FUNCTION_BLOCK basicGeradorGenerico (* Logica unica do grupo gerador (DEIF AGC 150): valores, estado do QTA, modo e alarmes *)
  (* Standard: 61499-2 *)
  (* Version 1.1, 15/10/2026, Hidryco, Hidryco, 1.1: comandos basicos (automatico, semiautomatico, partir, parar, reconhecer alarmes do AGC) nas palavras 5 e 6. 1.0: AGC 150 (GEN) por Modbus TCP FC04, tabela DEIF rev. S; so supervisao *)
  PACKAGE Hidryco.HidrycoLib;
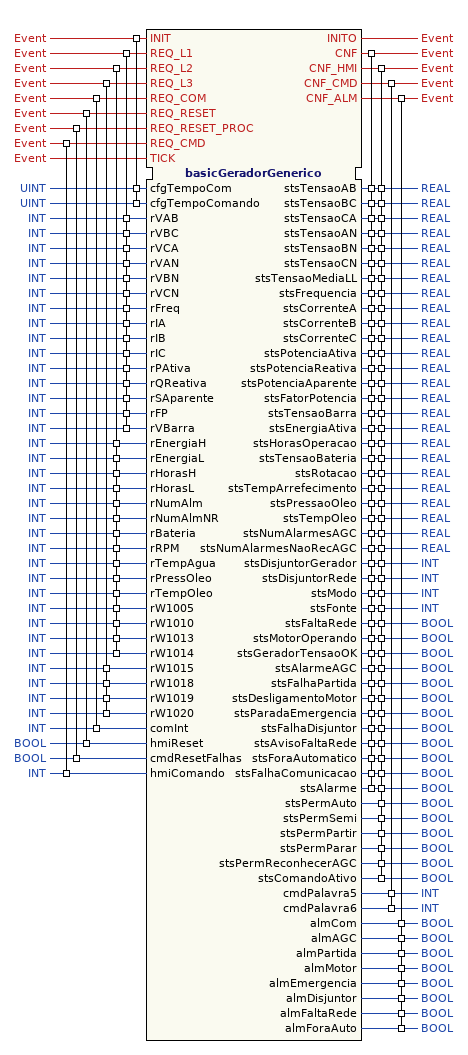
  EVENT_INPUT
    INIT WITH cfgTempoCom, cfgTempoComando; (* Inicializacao *)
    REQ_L1 WITH rVAB, rVBC, rVCA, rVAN, rVBN, rVCN, rFreq, rIA, rIB, rIC, rPAtiva, rQReativa, rSAparente, rFP, rVBarra; (* Leitura 1 (grandezas eletricas) *)
    REQ_L2 WITH rEnergiaH, rEnergiaL, rHorasH, rHorasL, rNumAlm, rNumAlmNR, rBateria, rRPM, rTempAgua, rPressOleo, rTempOleo, rW1005, rW1010, rW1013, rW1014; (* Leitura 2 (contadores, motor, alarmes) *)
    REQ_L3 WITH rW1015, rW1018, rW1019, rW1020; (* Leitura 3 (estado e modos) *)
    REQ_COM WITH comInt; (* Comunicacao *)
    REQ_RESET WITH hmiReset; (* Reconhecimento pela IHM *)
    REQ_RESET_PROC WITH cmdResetFalhas; (* Reconhecimento pelo processo *)
    REQ_CMD WITH hmiComando; (* Comando da IHM para o AGC *)
    TICK; (* Base de tempo de 1 s (E_CYCLE) *)
  END_EVENT
  EVENT_OUTPUT
    INITO; (* Inicializacao concluida *)
    CNF WITH stsTensaoAB, stsTensaoBC, stsTensaoCA, stsTensaoAN, stsTensaoBN, stsTensaoCN, stsTensaoMediaLL, stsFrequencia, stsCorrenteA, stsCorrenteB, stsCorrenteC, stsPotenciaAtiva, stsPotenciaReativa, stsPotenciaAparente, stsFatorPotencia, stsTensaoBarra, stsEnergiaAtiva, stsHorasOperacao, stsTensaoBateria, stsRotacao, stsTempArrefecimento, stsPressaoOleo, stsTempOleo, stsNumAlarmesAGC, stsNumAlarmesNaoRecAGC, stsDisjuntorGerador, stsDisjuntorRede, stsModo, stsFonte, stsFaltaRede, stsMotorOperando, stsGeradorTensaoOK, stsAlarmeAGC, stsFalhaPartida, stsDesligamentoMotor, stsParadaEmergencia, stsFalhaDisjuntor, stsAvisoFaltaRede, stsForaAutomatico, stsFalhaComunicacao, stsAlarme; (* Valores e estados (na mudanca) *)
    CNF_HMI WITH stsTensaoAB, stsTensaoBC, stsTensaoCA, stsTensaoAN, stsTensaoBN, stsTensaoCN, stsTensaoMediaLL, stsFrequencia, stsCorrenteA, stsCorrenteB, stsCorrenteC, stsPotenciaAtiva, stsPotenciaReativa, stsPotenciaAparente, stsFatorPotencia, stsTensaoBarra, stsEnergiaAtiva, stsHorasOperacao, stsTensaoBateria, stsRotacao, stsTempArrefecimento, stsPressaoOleo, stsTempOleo, stsNumAlarmesAGC, stsNumAlarmesNaoRecAGC, stsDisjuntorGerador, stsDisjuntorRede, stsModo, stsFonte, stsFaltaRede, stsMotorOperando, stsGeradorTensaoOK, stsAlarmeAGC, stsFalhaPartida, stsDesligamentoMotor, stsParadaEmergencia, stsFalhaDisjuntor, stsAvisoFaltaRede, stsForaAutomatico, stsFalhaComunicacao, stsAlarme, stsPermAuto, stsPermSemi, stsPermPartir, stsPermParar, stsPermReconhecerAGC, stsComandoAtivo; (* Status para a IHM (na mudanca) *)
    CNF_CMD WITH cmdPalavra5, cmdPalavra6; (* Palavras de comando do AGC (na mudanca) *)
    CNF_ALM WITH almCom, almAGC, almPartida, almMotor, almEmergencia, almDisjuntor, almFaltaRede, almForaAuto; (* Alarmes para os ALARM_BIT (na mudanca) *)
  END_EVENT
  VAR_INPUT
    cfgTempoCom : UINT := 10; (* Tempo (s) sem comunicacao com o AGC 150 para confirmar a falha *)
    cfgTempoComando : UINT := 2; (* Tempo (s) que a palavra de comando fica escrita no AGC *)
    rVAB : INT; (* Tensao do gerador L1-L2 (V) *)
    rVBC : INT; (* Tensao do gerador L2-L3 (V) *)
    rVCA : INT; (* Tensao do gerador L3-L1 (V) *)
    rVAN : INT; (* Tensao do gerador L1-N (V) *)
    rVBN : INT; (* Tensao do gerador L2-N (V) *)
    rVCN : INT; (* Tensao do gerador L3-N (V) *)
    rFreq : INT; (* Frequencia do gerador L1 (0,01 Hz) *)
    rIA : INT; (* Corrente do gerador L1 (A) *)
    rIB : INT; (* Corrente do gerador L2 (A) *)
    rIC : INT; (* Corrente do gerador L3 (A) *)
    rPAtiva : INT; (* Potencia ativa do gerador (kW) *)
    rQReativa : INT; (* Potencia reativa do gerador (kVAr) *)
    rSAparente : INT; (* Potencia aparente do gerador (kVA) *)
    rFP : INT; (* Fator de potencia do gerador (0,01) *)
    rVBarra : INT; (* Tensao do lado B (barramento/rede) L1-L2 (V) *)
    rEnergiaH : INT; (* Energia ativa exportada total - palavra alta (INT32 ABCD, kWh) *)
    rEnergiaL : INT; (* Energia ativa exportada total - palavra baixa *)
    rHorasH : INT; (* Horas de funcionamento absolutas - palavra alta (INT32 ABCD, h) *)
    rHorasL : INT; (* Horas de funcionamento absolutas - palavra baixa *)
    rNumAlm : INT; (* Numero de alarmes ativos no AGC *)
    rNumAlmNR : INT; (* Numero de alarmes nao reconhecidos no AGC *)
    rBateria : INT; (* Tensao de alimentacao DC (bateria), term. 1-2 (0,1 V) *)
    rRPM : INT; (* Rotacao do motor - ECU (rpm) *)
    rTempAgua : INT; (* Temperatura do liquido de arrefecimento - ECU (0,1 C) *)
    rPressOleo : INT; (* Pressao do oleo - ECU (0,01 bar) *)
    rTempOleo : INT; (* Temperatura do oleo - ECU (0,1 C) *)
    rW1005 : INT; (* Alarmes de disjuntor e sincronismo (bits) *)
    rW1010 : INT; (* Alarmes de entradas digitais (bit 12 = parada de emergencia) *)
    rW1013 : INT; (* Alarmes do motor (bits: 9/10 sobrevelocidade, 11 falha de arranque, 15 falha de partida) *)
    rW1014 : INT; (* Alarmes do motor (bit 0 = falha de parada) *)
    rW1015 : INT; (* Alarmes diversos (bit 12 = fora do automatico) *)
    rW1018 : INT; (* Estado da planta (bits: 0 falta de rede, 1 MB ON, 4 GB ON, 6 motor em operacao, 8 Hz/V OK, 11 GB OFF, 12 MB OFF) *)
    rW1019 : INT; (* Modos (bits: 0 bloqueio, 1 manual, 2 semi-auto, 3 auto, 4 teste) *)
    rW1020 : INT; (* Alarmes da ECU (bit 2 = shutdown / alarme vermelho) *)
    comInt : INT; (* connStatusInt do MODBUSGENTCPS (1 = online) *)
    hmiReset : BOOL; (* IHM: reconhecimento *)
    cmdResetFalhas : BOOL; (* Processo: reconhecimento (com E_RESET_FALHAS) *)
    hmiComando : INT; (* IHM: comando para o AGC (1 automatico, 2 semiautomatico, 3 partir, 4 parar, 5 reconhecer alarmes do AGC) *)
  END_VAR
  VAR_OUTPUT
    stsTensaoAB : REAL; (* Tensao A-B (V) *)
    stsTensaoBC : REAL; (* Tensao B-C (V) *)
    stsTensaoCA : REAL; (* Tensao C-A (V) *)
    stsTensaoAN : REAL; (* Tensao A-N (V) *)
    stsTensaoBN : REAL; (* Tensao B-N (V) *)
    stsTensaoCN : REAL; (* Tensao C-N (V) *)
    stsTensaoMediaLL : REAL; (* Tensao media fase-fase (V) *)
    stsFrequencia : REAL; (* Frequencia (Hz) *)
    stsCorrenteA : REAL; (* Corrente fase A (A) *)
    stsCorrenteB : REAL; (* Corrente fase B (A) *)
    stsCorrenteC : REAL; (* Corrente fase C (A) *)
    stsPotenciaAtiva : REAL; (* Potencia ativa (kW) *)
    stsPotenciaReativa : REAL; (* Potencia reativa (kVAr) *)
    stsPotenciaAparente : REAL; (* Potencia aparente (kVA) *)
    stsFatorPotencia : REAL; (* Fator de potencia *)
    stsTensaoBarra : REAL; (* Tensao do lado B (barramento/rede) L1-L2 (V) *)
    stsEnergiaAtiva : REAL; (* Energia ativa exportada (kWh) *)
    stsHorasOperacao : REAL; (* Horas de funcionamento (h) *)
    stsTensaoBateria : REAL; (* Tensao da bateria (V) *)
    stsRotacao : REAL; (* Rotacao do motor (rpm) *)
    stsTempArrefecimento : REAL; (* Temperatura do liquido de arrefecimento (°C) *)
    stsPressaoOleo : REAL; (* Pressao do oleo (bar) *)
    stsTempOleo : REAL; (* Temperatura do oleo (°C) *)
    stsNumAlarmesAGC : REAL; (* Alarmes ativos no AGC *)
    stsNumAlarmesNaoRecAGC : REAL; (* Alarmes nao reconhecidos no AGC *)
    stsDisjuntorGerador : INT; (* Disjuntor do gerador (GB): 0 indefinido/sem comunicacao, 1 aberto, 2 fechado *)
    stsDisjuntorRede : INT; (* Disjuntor de rede (MB): 0 indefinido/sem comunicacao, 1 aberto, 2 fechado *)
    stsModo : INT; (* Modo do AGC: 0 indefinido, 1 automatico, 2 semi-automatico, 3 manual, 4 bloqueio, 5 teste *)
    stsFonte : INT; (* Fonte da saida do QTA: 0 sem fonte, 1 rede, 2 gerador, 3 indefinida (sem comunicacao) *)
    stsFaltaRede : BOOL; (* Falta de rede (AMF) *)
    stsMotorOperando : BOOL; (* Motor em operacao *)
    stsGeradorTensaoOK : BOOL; (* Tensao e frequencia do gerador OK *)
    stsAlarmeAGC : BOOL; (* Alarme ativo no controlador do gerador (AGC 150) *)
    stsFalhaPartida : BOOL; (* Falha na partida do gerador *)
    stsDesligamentoMotor : BOOL; (* Desligamento do motor (ECU ou sobrevelocidade) *)
    stsParadaEmergencia : BOOL; (* Parada de emergência do gerador acionada *)
    stsFalhaDisjuntor : BOOL; (* Falha de disjuntor no QTA (gerador ou rede) *)
    stsAvisoFaltaRede : BOOL; (* Falta de rede no QTA *)
    stsForaAutomatico : BOOL; (* Gerador fora do modo automático *)
    stsFalhaComunicacao : BOOL; (* Falha de comunicacao com o AGC 150 *)
    stsAlarme : BOOL; (* Algum alarme do gerador *)
    stsPermAuto : BOOL; (* IHM: comando Auto permitido *)
    stsPermSemi : BOOL; (* IHM: comando Semi permitido *)
    stsPermPartir : BOOL; (* IHM: comando Partir permitido *)
    stsPermParar : BOOL; (* IHM: comando Parar permitido *)
    stsPermReconhecerAGC : BOOL; (* IHM: comando ReconhecerAGC permitido *)
    stsComandoAtivo : BOOL; (* Comando sendo enviado ao AGC *)
    cmdPalavra5 : INT; (* Palavra de comando 5 do AGC (holding register 5) *)
    cmdPalavra6 : INT; (* Palavra de comando 6 do AGC (holding register 6) *)
    almCom : BOOL; (* ALARM_BIT falha de comunicacao *)
    almAGC : BOOL; (* ALARM_BIT Alarme ativo no controlador do gerador (AGC 150) *)
    almPartida : BOOL; (* ALARM_BIT Falha na partida do gerador *)
    almMotor : BOOL; (* ALARM_BIT Desligamento do motor (ECU ou sobrevelocidade) *)
    almEmergencia : BOOL; (* ALARM_BIT Parada de emergência do gerador acionada *)
    almDisjuntor : BOOL; (* ALARM_BIT Falha de disjuntor no QTA (gerador ou rede) *)
    almFaltaRede : BOOL; (* ALARM_BIT Falta de rede no QTA *)
    almForaAuto : BOOL; (* ALARM_BIT Gerador fora do modo automático *)
  END_VAR
  VAR
    initDone : BOOL;
    initPass : BOOL;
    bComRecebida : BOOL; (* Ja houve leitura do connStatusInt *)
    bValido : BOOL; (* AGC comunicando: valores validos *)
    uSegCom : UDINT;
    w05 : WORD;
    w10 : WORD;
    w13 : WORD;
    w18 : WORD;
    w19 : WORD;
    w20 : WORD;
    bGBon : BOOL;
    bGBoff : BOOL;
    bMBon : BOOL;
    bMBoff : BOOL;
    bMudou : BOOL;
    wSts : DWORD;
    oldSts : DWORD := 16#FFFFFFFF;
    wAlm : WORD;
    oldAlm : WORD := 16#FFFF;
    iOld : INT;
    uCmd : UINT; (* Segundos restantes do pulso de comando *)
    wPerm : WORD;
    oldPerm : WORD := 16#FFFF;
    o_stsTensaoAB : REAL := -1.0;
    o_stsTensaoBC : REAL := -1.0;
    o_stsTensaoCA : REAL := -1.0;
    o_stsTensaoAN : REAL := -1.0;
    o_stsTensaoBN : REAL := -1.0;
    o_stsTensaoCN : REAL := -1.0;
    o_stsTensaoMediaLL : REAL := -1.0;
    o_stsFrequencia : REAL := -1.0;
    o_stsCorrenteA : REAL := -1.0;
    o_stsCorrenteB : REAL := -1.0;
    o_stsCorrenteC : REAL := -1.0;
    o_stsPotenciaAtiva : REAL := -1.0;
    o_stsPotenciaReativa : REAL := -1.0;
    o_stsPotenciaAparente : REAL := -1.0;
    o_stsFatorPotencia : REAL := -1.0;
    o_stsTensaoBarra : REAL := -1.0;
    o_stsEnergiaAtiva : REAL := -1.0;
    o_stsHorasOperacao : REAL := -1.0;
    o_stsTensaoBateria : REAL := -1.0;
    o_stsRotacao : REAL := -1.0;
    o_stsTempArrefecimento : REAL := -1.0;
    o_stsPressaoOleo : REAL := -1.0;
    o_stsTempOleo : REAL := -1.0;
    o_stsNumAlarmesAGC : REAL := -1.0;
    o_stsNumAlarmesNaoRecAGC : REAL := -1.0;
    o_stsDisjuntorGerador : INT := -1;
    o_stsDisjuntorRede : INT := -1;
    o_stsModo : INT := -1;
    o_stsFonte : INT := -1;
  END_VAR
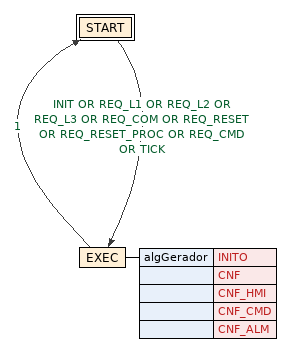
  EC_STATES
    START; (* Estado inicial *)
    EXEC : algGerador -> INITO, -> CNF, -> CNF_HMI, -> CNF_CMD, -> CNF_ALM; (* Executa a logica; o algoritmo decide quais eventos saem *)
  END_STATES
  EC_TRANSITIONS
    START TO EXEC := INIT OR REQ_L1 OR REQ_L2 OR REQ_L3 OR REQ_COM OR REQ_RESET OR REQ_RESET_PROC OR REQ_CMD OR TICK;
    EXEC TO START := 1;
  END_TRANSITIONS
  ALGORITHM algGerador IN ST: (* Logica completa do gerador (um unico algoritmo) *)
(* =====================================================================
   basicGeradorGenerico v1.0 - grupo gerador com controlador DEIF AGC 150
   (aplicacao GEN: QTA com disjuntor do gerador GB e de rede MB)
   Registradores de entrada (FC04) da tabela DEIF "AGC 150 Modbus server
   tables" rev. S (software 1.19). v1.1: comandos basicos nas palavras de
   comando 5 e 6 (pulso de cfgTempoComando s; depois as palavras voltam a 0).
   Padrao das bibliotecas Schneider: eventos de saida desligados no inicio e
   ligados so na mudanca; tempos contados pelo TICK de 1 s (E_CYCLE do CAT).
   - escalas da tabela: frequencia e FP 0,01; bateria, temperaturas 0,1;
     pressao do oleo 0,01 bar; energia e horas INT32 (ABCD, palavra alta 1o);
   - falha de comunicacao: connStatusInt <> 1 por cfgTempoCom s; com a
     falha os estados ficam indefinidos e os demais alarmes suprimidos;
   - alarmes seguem o AGC (nao memorizados aqui): o reconhecimento na IHM
     reconhece os ALARM_BIT; os alarmes do AGC sao reconhecidos no AGC.
   ===================================================================== *)

INITO   := FALSE;
CNF     := FALSE;
CNF_HMI := FALSE;
CNF_CMD := FALSE;
CNF_ALM := FALSE;

IF REQ_COM THEN
    bComRecebida := TRUE;
END_IF;
IF INIT THEN
    initDone := TRUE;
    initPass := TRUE;
    INITO    := TRUE;
END_IF;
IF NOT initDone THEN
    RETURN;
END_IF;

(* ---- 1. Comunicacao ---- *)
IF comInt <> 1 THEN
    IF TICK AND uSegCom < UINT_TO_UDINT(cfgTempoCom) THEN
        uSegCom := uSegCom + 1;
    END_IF;
ELSE
    uSegCom := 0;
END_IF;
stsFalhaComunicacao := comInt <> 1 AND uSegCom >= UINT_TO_UDINT(cfgTempoCom);
bValido := bComRecebida AND comInt = 1;

(* ---- 2. Valores (ficam congelados sem comunicacao) ---- *)
stsTensaoAB := INT_TO_REAL(rVAB);
stsTensaoBC := INT_TO_REAL(rVBC);
stsTensaoCA := INT_TO_REAL(rVCA);
stsTensaoAN := INT_TO_REAL(rVAN);
stsTensaoBN := INT_TO_REAL(rVBN);
stsTensaoCN := INT_TO_REAL(rVCN);
stsTensaoMediaLL := (INT_TO_REAL(rVAB) + INT_TO_REAL(rVBC) + INT_TO_REAL(rVCA)) / 3.0;
stsFrequencia := INT_TO_REAL(rFreq) / 100.0;
stsCorrenteA := INT_TO_REAL(rIA);
stsCorrenteB := INT_TO_REAL(rIB);
stsCorrenteC := INT_TO_REAL(rIC);
stsPotenciaAtiva := INT_TO_REAL(rPAtiva);
stsPotenciaReativa := INT_TO_REAL(rQReativa);
stsPotenciaAparente := INT_TO_REAL(rSAparente);
stsFatorPotencia := INT_TO_REAL(rFP) / 100.0;
stsTensaoBarra := INT_TO_REAL(rVBarra);
stsEnergiaAtiva := DINT_TO_REAL(DWORD_TO_DINT(SHL(WORD_TO_DWORD(INT_TO_WORD(rEnergiaH)), 16) OR WORD_TO_DWORD(INT_TO_WORD(rEnergiaL))));
stsHorasOperacao := DINT_TO_REAL(DWORD_TO_DINT(SHL(WORD_TO_DWORD(INT_TO_WORD(rHorasH)), 16) OR WORD_TO_DWORD(INT_TO_WORD(rHorasL))));
stsTensaoBateria := INT_TO_REAL(rBateria) / 10.0;
stsRotacao := INT_TO_REAL(rRPM);
stsTempArrefecimento := INT_TO_REAL(rTempAgua) / 10.0;
stsPressaoOleo := INT_TO_REAL(rPressOleo) / 100.0;
stsTempOleo := INT_TO_REAL(rTempOleo) / 10.0;
stsNumAlarmesAGC := INT_TO_REAL(rNumAlm);
stsNumAlarmesNaoRecAGC := INT_TO_REAL(rNumAlmNR);

(* ---- 3. Palavras de estado e alarme ---- *)
w05 := INT_TO_WORD(rW1005);
w10 := INT_TO_WORD(rW1010);
w13 := INT_TO_WORD(rW1013);
w18 := INT_TO_WORD(rW1018);
w19 := INT_TO_WORD(rW1019);
w20 := INT_TO_WORD(rW1020);
bGBon  := (w18 AND 16#0010) <> 16#0000;
bGBoff := (w18 AND 16#0800) <> 16#0000;
bMBon  := (w18 AND 16#0002) <> 16#0000;
bMBoff := (w18 AND 16#1000) <> 16#0000;

stsFaltaRede := bValido AND ((w18 AND 16#0001) <> 16#0000);
stsMotorOperando := bValido AND ((w18 AND 16#0040) <> 16#0000);
stsGeradorTensaoOK := bValido AND ((w18 AND 16#0100) <> 16#0000);

(* disjuntores: 2 fechado, 1 aberto, 0 indefinido (transicao ou sem comunicacao) *)
IF NOT bValido THEN
    stsDisjuntorGerador := 0;
    stsDisjuntorRede := 0;
ELSE
    IF bGBon AND NOT bGBoff THEN stsDisjuntorGerador := 2;
    ELSIF bGBoff AND NOT bGBon THEN stsDisjuntorGerador := 1;
    ELSE stsDisjuntorGerador := 0;
    END_IF;
    IF bMBon AND NOT bMBoff THEN stsDisjuntorRede := 2;
    ELSIF bMBoff AND NOT bMBon THEN stsDisjuntorRede := 1;
    ELSE stsDisjuntorRede := 0;
    END_IF;
END_IF;

(* modo: teste > bloqueio > manual > semi > auto *)
IF NOT bValido THEN stsModo := 0;
ELSIF (w19 AND 16#0010) <> 16#0000 THEN stsModo := 5;
ELSIF (w19 AND 16#0001) <> 16#0000 THEN stsModo := 4;
ELSIF (w19 AND 16#0002) <> 16#0000 THEN stsModo := 3;
ELSIF (w19 AND 16#0004) <> 16#0000 THEN stsModo := 2;
ELSIF (w19 AND 16#0008) <> 16#0000 THEN stsModo := 1;
ELSE stsModo := 0;
END_IF;

(* fonte da saida do QTA *)
IF NOT bValido THEN stsFonte := 3;
ELSIF stsDisjuntorGerador = 2 THEN stsFonte := 2;
ELSIF stsDisjuntorRede = 2 THEN stsFonte := 1;
ELSE stsFonte := 0;
END_IF;

(* ---- 4. Alarmes (seguem o AGC; so com comunicacao) ---- *)
stsAlarmeAGC := bValido AND (rNumAlm > 0);
stsFalhaPartida := bValido AND ((w13 AND 16#8800) <> 16#0000);
stsDesligamentoMotor := bValido AND (((w20 AND 16#0004) <> 16#0000) OR ((w13 AND 16#0600) <> 16#0000));
stsParadaEmergencia := bValido AND ((w10 AND 16#1000) <> 16#0000);
stsFalhaDisjuntor := bValido AND ((w05 AND 16#03F0) <> 16#0000);
stsAvisoFaltaRede := bValido AND ((w18 AND 16#0001) <> 16#0000);
stsForaAutomatico := bValido AND ((w19 AND 16#0008) = 16#0000);

almCom := stsFalhaComunicacao;
almAGC := stsAlarmeAGC;
almPartida := stsFalhaPartida;
almMotor := stsDesligamentoMotor;
almEmergencia := stsParadaEmergencia;
almDisjuntor := stsFalhaDisjuntor;
almFaltaRede := stsAvisoFaltaRede;
almForaAuto := stsForaAutomatico;
stsAlarme := almCom OR almAGC OR almPartida OR almMotor OR almEmergencia OR almDisjuntor OR almFaltaRede OR almForaAuto;

(* ---- 5. Comandos basicos (IHM) nas palavras 5 e 6 do AGC ---- *)
stsPermAuto := bValido AND stsModo <> 1;
stsPermSemi := bValido AND stsModo <> 2;
stsPermPartir := bValido AND stsModo = 2 AND NOT stsMotorOperando;
stsPermParar := bValido AND stsModo = 2 AND stsMotorOperando;
stsPermReconhecerAGC := bValido;
IF REQ_CMD AND uCmd = 0 THEN
    IF hmiComando = 1 AND stsPermAuto THEN
        cmdPalavra6 := 8193; cmdPalavra5 := 0;
        uCmd := cfgTempoComando + 1;
        CNF_CMD := TRUE;
    ELSIF hmiComando = 2 AND stsPermSemi THEN
        cmdPalavra6 := 16385; cmdPalavra5 := 0;
        uCmd := cfgTempoComando + 1;
        CNF_CMD := TRUE;
    ELSIF hmiComando = 3 AND stsPermPartir THEN
        cmdPalavra5 := 3; cmdPalavra6 := 0;
        uCmd := cfgTempoComando + 1;
        CNF_CMD := TRUE;
    ELSIF hmiComando = 4 AND stsPermParar THEN
        cmdPalavra5 := 17; cmdPalavra6 := 0;
        uCmd := cfgTempoComando + 1;
        CNF_CMD := TRUE;
    ELSIF hmiComando = 5 AND stsPermReconhecerAGC THEN
        cmdPalavra5 := 1025; cmdPalavra6 := 0;
        uCmd := cfgTempoComando + 1;
        CNF_CMD := TRUE;
    END_IF;
END_IF;
IF TICK AND uCmd > 0 THEN
    uCmd := uCmd - 1;
    IF uCmd = 0 THEN
        cmdPalavra5 := 0;
        cmdPalavra6 := 0;
        CNF_CMD := TRUE;
    END_IF;
END_IF;
IF NOT bValido AND uCmd > 0 THEN
    uCmd := 0;
    cmdPalavra5 := 0;
    cmdPalavra6 := 0;
    CNF_CMD := TRUE;
END_IF;
stsComandoAtivo := uCmd > 0;
wPerm := 0;
IF stsPermAuto THEN wPerm := wPerm OR 16#0001; END_IF;
IF stsPermSemi THEN wPerm := wPerm OR 16#0002; END_IF;
IF stsPermPartir THEN wPerm := wPerm OR 16#0004; END_IF;
IF stsPermParar THEN wPerm := wPerm OR 16#0008; END_IF;
IF stsPermReconhecerAGC THEN wPerm := wPerm OR 16#0010; END_IF;
IF stsComandoAtivo THEN wPerm := wPerm OR 16#0020; END_IF;

(* ---- 6. Eventos so na mudanca ---- *)
bMudou := FALSE;
IF stsTensaoAB <> o_stsTensaoAB THEN bMudou := TRUE; o_stsTensaoAB := stsTensaoAB; END_IF;
IF stsTensaoBC <> o_stsTensaoBC THEN bMudou := TRUE; o_stsTensaoBC := stsTensaoBC; END_IF;
IF stsTensaoCA <> o_stsTensaoCA THEN bMudou := TRUE; o_stsTensaoCA := stsTensaoCA; END_IF;
IF stsTensaoAN <> o_stsTensaoAN THEN bMudou := TRUE; o_stsTensaoAN := stsTensaoAN; END_IF;
IF stsTensaoBN <> o_stsTensaoBN THEN bMudou := TRUE; o_stsTensaoBN := stsTensaoBN; END_IF;
IF stsTensaoCN <> o_stsTensaoCN THEN bMudou := TRUE; o_stsTensaoCN := stsTensaoCN; END_IF;
IF stsTensaoMediaLL <> o_stsTensaoMediaLL THEN bMudou := TRUE; o_stsTensaoMediaLL := stsTensaoMediaLL; END_IF;
IF stsFrequencia <> o_stsFrequencia THEN bMudou := TRUE; o_stsFrequencia := stsFrequencia; END_IF;
IF stsCorrenteA <> o_stsCorrenteA THEN bMudou := TRUE; o_stsCorrenteA := stsCorrenteA; END_IF;
IF stsCorrenteB <> o_stsCorrenteB THEN bMudou := TRUE; o_stsCorrenteB := stsCorrenteB; END_IF;
IF stsCorrenteC <> o_stsCorrenteC THEN bMudou := TRUE; o_stsCorrenteC := stsCorrenteC; END_IF;
IF stsPotenciaAtiva <> o_stsPotenciaAtiva THEN bMudou := TRUE; o_stsPotenciaAtiva := stsPotenciaAtiva; END_IF;
IF stsPotenciaReativa <> o_stsPotenciaReativa THEN bMudou := TRUE; o_stsPotenciaReativa := stsPotenciaReativa; END_IF;
IF stsPotenciaAparente <> o_stsPotenciaAparente THEN bMudou := TRUE; o_stsPotenciaAparente := stsPotenciaAparente; END_IF;
IF stsFatorPotencia <> o_stsFatorPotencia THEN bMudou := TRUE; o_stsFatorPotencia := stsFatorPotencia; END_IF;
IF stsTensaoBarra <> o_stsTensaoBarra THEN bMudou := TRUE; o_stsTensaoBarra := stsTensaoBarra; END_IF;
IF stsEnergiaAtiva <> o_stsEnergiaAtiva THEN bMudou := TRUE; o_stsEnergiaAtiva := stsEnergiaAtiva; END_IF;
IF stsHorasOperacao <> o_stsHorasOperacao THEN bMudou := TRUE; o_stsHorasOperacao := stsHorasOperacao; END_IF;
IF stsTensaoBateria <> o_stsTensaoBateria THEN bMudou := TRUE; o_stsTensaoBateria := stsTensaoBateria; END_IF;
IF stsRotacao <> o_stsRotacao THEN bMudou := TRUE; o_stsRotacao := stsRotacao; END_IF;
IF stsTempArrefecimento <> o_stsTempArrefecimento THEN bMudou := TRUE; o_stsTempArrefecimento := stsTempArrefecimento; END_IF;
IF stsPressaoOleo <> o_stsPressaoOleo THEN bMudou := TRUE; o_stsPressaoOleo := stsPressaoOleo; END_IF;
IF stsTempOleo <> o_stsTempOleo THEN bMudou := TRUE; o_stsTempOleo := stsTempOleo; END_IF;
IF stsNumAlarmesAGC <> o_stsNumAlarmesAGC THEN bMudou := TRUE; o_stsNumAlarmesAGC := stsNumAlarmesAGC; END_IF;
IF stsNumAlarmesNaoRecAGC <> o_stsNumAlarmesNaoRecAGC THEN bMudou := TRUE; o_stsNumAlarmesNaoRecAGC := stsNumAlarmesNaoRecAGC; END_IF;
IF stsDisjuntorGerador <> o_stsDisjuntorGerador THEN bMudou := TRUE; o_stsDisjuntorGerador := stsDisjuntorGerador; END_IF;
IF stsDisjuntorRede <> o_stsDisjuntorRede THEN bMudou := TRUE; o_stsDisjuntorRede := stsDisjuntorRede; END_IF;
IF stsModo <> o_stsModo THEN bMudou := TRUE; o_stsModo := stsModo; END_IF;
IF stsFonte <> o_stsFonte THEN bMudou := TRUE; o_stsFonte := stsFonte; END_IF;
wSts := 0;
IF stsFaltaRede THEN wSts := wSts OR 16#00000001; END_IF;
IF stsMotorOperando THEN wSts := wSts OR 16#00000002; END_IF;
IF stsGeradorTensaoOK THEN wSts := wSts OR 16#00000004; END_IF;
IF stsAlarmeAGC THEN wSts := wSts OR 16#00000008; END_IF;
IF stsFalhaPartida THEN wSts := wSts OR 16#00000010; END_IF;
IF stsDesligamentoMotor THEN wSts := wSts OR 16#00000020; END_IF;
IF stsParadaEmergencia THEN wSts := wSts OR 16#00000040; END_IF;
IF stsFalhaDisjuntor THEN wSts := wSts OR 16#00000080; END_IF;
IF stsAvisoFaltaRede THEN wSts := wSts OR 16#00000100; END_IF;
IF stsForaAutomatico THEN wSts := wSts OR 16#00000200; END_IF;
IF stsFalhaComunicacao THEN wSts := wSts OR 16#00000400; END_IF;
IF stsAlarme THEN wSts := wSts OR 16#00000800; END_IF;
wAlm := 0;
IF almCom THEN wAlm := wAlm OR 16#0001; END_IF;
IF almAGC THEN wAlm := wAlm OR 16#0002; END_IF;
IF almPartida THEN wAlm := wAlm OR 16#0004; END_IF;
IF almMotor THEN wAlm := wAlm OR 16#0008; END_IF;
IF almEmergencia THEN wAlm := wAlm OR 16#0010; END_IF;
IF almDisjuntor THEN wAlm := wAlm OR 16#0020; END_IF;
IF almFaltaRede THEN wAlm := wAlm OR 16#0040; END_IF;
IF almForaAuto THEN wAlm := wAlm OR 16#0080; END_IF;
CNF := initPass OR bMudou OR (wSts <> oldSts);
CNF_HMI := CNF OR (wPerm <> oldPerm);
IF initPass THEN
    CNF_CMD := TRUE;
END_IF;
CNF_ALM := initPass OR (wAlm <> oldAlm);
oldSts := wSts;
oldPerm := wPerm;
oldAlm := wAlm;
initPass := FALSE;
  END_ALGORITHM
END_FUNCTION_BLOCK
